TYPE "ST_CylinderOutCmd"
VERSION : 0.1
   STRUCT
      Direction : DInt;
   END_STRUCT;

END_TYPE

